Fanuc KAREL source: kc00034.KL

-- PROVISIONAL review KL for V1013-1; original PC SHA256 e0388d21fcfcad248aca539a48d207cca2ac53c6e3e8d4f38f30b9c4d041ffe9
-- Incomplete behavior may be omitted. Consult companion uncertainty JSON. Do not deploy.
PROGRAM KC00034
%NOLOCKGROUP
BEGIN
  -- UNRESOLVED_PC offsets 5-29; opcodes 27,22,22,2A,22,31
  -- UNRESOLVED_PC offsets 34-38; opcodes 7F
END KC00034
